Staubli VAL3: exercice6.pgx

program exercice6()
  local num l_nNbKapla
  local pointRx dest
  local trsf Pas
  local trsf Decal
begin

  wait(bInit_repere == true)
  for l_nNbKapla = 0 to 4

    Decal.x = l_nNbKapla * 40

    dest = compose(plA,fcaisse,Decal)

    bStart = false
    nCouleur_Autorisation = "#80EA34"
    movej(appro(dest,{0,0,-50,0,0,0}),tPince,mRapide)
    movel(dest,tPince,mLent)
    call fermerPince()
    movel(appro(dest,{0,0,-50,0,0,0}),tPince,mRapide)
    movej(jDepart,tPince,mRapide)

    wait(bStart == true)
    nCouleur_Autorisation = "#EA3734"
    movej(appro(pDepose[0],{0,0,-50,0,0,0}),tPince,mRapide)
    movel(pDepose[0],tPince,mLent)
    call ouvrirPince()
    movel(appro(pDepose[0],{0,0,-50,0,0,0}),tPince,mRapide)
    movej(jDepart,tPince,mLent)
    waitEndMove()


  endFor
end
